TYPE str_ConcParam :
	//to be deletd
STRUCT
	
    r_Temper_1			:	REAL:=65	;//temperature set point for local client in celsius
	r_Flow_Pmp1_1		:	REAL:=180	;
	r_Flow_Pmp1_2		:	REAL:=180	;
	r_Pressure_Pmp1_1	:	REAL:=0.5	;
	r_Concentration_1	:	REAL:=0.3	;//concentration in percents
	t_Measure_Delay_1	:	INT:=60		;//measurment delay in seconds
END_STRUCT
END_TYPE

(* stored: Version 1.1.0.1, ProductVersion 3.1.4024.12
   DUT str_ConcParam: Id {50f78a7b-79b6-4e73-81c5-8e0b587658a9} *)
